// TIA Portal V14 SP1 export
// export: Created 2000-01-01T00:00:00.0000000Z, ExportSetting None
DATA_BLOCK "MCP_RC_DB2"   // DB9802
{ S7_Optimized_Access := 'TRUE' }
   VAR
      Count : Int := 4;
      Motor : "MCP_RC_UDT";
   END_VAR
BEGIN
   Motor.Speed := 11;
END_DATA_BLOCK
